(* IEC 61131-3 sources: axsharp/src/ix.templates/working/templates/ixblazor/ax/src, 3 files *)

(* ---- counters.st ---- *)
CLASS Counters
    VAR PUBLIC
        {#ix-attr:[Container(Layout.Wrap)]}
        wrap : Counter;
        {#ix-attr:[Container(Layout.Stack)]}
        stack : Counter;
        {#ix-attr:[Container(Layout.UniformGrid)]}
        grid : Counter;
        {#ix-attr:[Container(Layout.Tabs)]}
        tabs : Counter;
    END_VAR
END_CLASS

CLASS PUBLIC Counter
    VAR PUBLIC
        {#ix-set:AttributeName = "Number of revolutions"}
        Counts : ULINT;
        {#ix-set:AttributeName = "Count revolutions"}
        AllowCounter : BOOL;
        {#ix-set:AttributeName = "Reset counts"}
        ResetCounter : BOOL;
    END_VAR

    METHOD PUBLIC RunCounter
        IF (AllowCounter) THEN
            Counts := Counts + ULINT#1;
        END_IF;

        IF(ResetCounter) THEN
            Counts := ULINT#0;
            ResetCounter := FALSE;
        END_IF;
    END_METHOD
END_CLASS

(* ---- configuration.st ---- *)
CONFIGURATION MyConfiguration
    TASK Main(Interval := T#10ms, Priority := 1);
    PROGRAM P1 WITH Main: MyProgram;

    VAR_GLOBAL
       counters : counters;
    END_VAR
END_CONFIGURATION

(* ---- program.st ---- *)
PROGRAM MyProgram
    VAR_EXTERNAL
        counters : counters;
    END_VAR
    counters.wrap.RunCounter();
    counters.stack.RunCounter();
    counters.grid.RunCounter();
    counters.tabs.RunCounter();
END_PROGRAM
